(* IEC 61131-3 sources: moqui-plc/codesys-v4/moqui-plc.fbsdev/moqui.iecapp^/moqui/framework/src/main/org/moqui/mqtt, 4 files *)

(* ---- MqttConnectionFactory.fb.st ---- *)
(* Component to connect with a MQTT broker, using default configurations. *)
FUNCTION_BLOCK MqttConnectionFactory

	VAR_INPUT
		connect : BOOL := TRUE;
	END_VAR
	VAR_OUTPUT
		connection : MQTT.MQTTClient;
	    connected : BOOL;
	    busy : BOOL;
	    error : BOOL;
		errorId : INT;
	END_VAR
	VAR
		(* Connect properties v5 *)
		mqttConnectProperties : MQTT.MQTTConnectProperties := (
			udiSessionExpiryInterval := MoquiConf.sessionExpiryInterval,
			udiMaximumPacketSize := MoquiConf.maximumPacketSize
			(* userProperties := connectUserProperties *)
		);
		(* Will properties v5 *)
		mqttWillProperties : MQTT.MQTTWillProperties := (
			bPayloadFormatIndicator := MoquiConf.willPayloadFormatIndicator,
			udiMessageExpiryInterval := MoquiConf.willMessageExpiryInterval,
			wsContentType := MoquiConf.willContentType,
			udiWillDelayInterval := MoquiConf.willDelayInterval
			(* userProperties := willUserProperties *)
	    );
		(* TLS context *)
		cipherList : NBS.CIPHER_LIST := (psList := ADR('HIGH'), udiSize := 5);
		commonName : STRING := 'moqui';
	    certInfo : NBS.CERT_INFO := (psInfo := ADR(commonName), udiSize := INT_TO_UDINT(LEN(commonName)));
		defaultTlsContext : NBS.TLSContext := (
			sUseCaseName := commonName,
			ePurpose := NBS.PURPOSE.CLIENT_SIDE,
			sTLSVersion := '1.3',
			sCipherList := cipherList,
			sHostname := MoquiConf.brokerUrl,
			ciCertInfo := certInfo,
			udiVerificationMode	:= 2, (* 1 => No peer verification, 2 => Active Peer verification *)
			itfCertVerifer := 0
		);
		nullTlsContext : NBS.ITLSContext := 0;
		tlsContext : NBS.ITLSContext;
		useTLS : BOOL := FALSE;

		(*
	     * To use client certificates, configure the connection via the TLS context.
		 * Example:
		 *      commonName : STRING := 'COMMON_NAME_OF_CERTIFICATE'; // CN of the certificate (common name).
		 *      cipherList : NBS.CIPHER_LIST := (psList := ADR('HIGH'), udiSize := 5); // Cipher string see https://www.openssl.org/docs/man1.1.1/man1/ciphers.html
		 *      certInfo : NBS.CERT_INFO := (psInfo := ADR(commonName), udiSize := SIZEOF(commonName)); // CN of the certificate (common name)
		 *      tlsContext : NBS.TLSContext := (
		 *          sUseCaseName := commonName, // A certificate is stored in the certificate store with the use case name.
		 *          ePurpose := NBS.PURPOSE.CLIENT_SIDE, // For client certificates set this to NBS.PURPOSE.CLIENT_SIDE
	     *          sTLSVersion := '1.3', // The TLS version
	     *          sCipherList := cipherList, // Set the cipher list
	     *          sHostname := brokerUrl, // The hostname of the broker
	     *          udiVerificationMode := 2, // 2 => Active Peer verification
	     *          ciCertInfo := certInfo, // Set the cert info
	     *          itfCertVerifer := 0); // 0 => No Verifier
		 *      client : MQTT.MQTTClient := (itfTLSCOntext := _tlsContext);
		 * Use the method TLSContext.SetInitialValue to set the context while runtime and set the context via the input itfTLSCOntext of the client FB.
		 *)
	END_VAR

	(* TLS selection *)
	tlsContext := nullTlsContext;
	IF useTLS THEN tlsContext := defaultTlsContext; END_IF;

	(* Configure the MQTT connection *)
	connection(xEnable := connect, xConnectedToBroker => connected, xError => error, eMQTTerror => errorId,
		sHostname := MoquiConf.brokerUrl, uiPort := MoquiConf.brokerPort, sWebSocketUrl := MoquiConf.webSocketUrl, sClientId := MoquiConf.clientId,
		itfTLSContext := tlsContext, eCommunicationMode := MoquiConf.communicationMode, eMQTTVersion := MoquiConf.mqttVersion,
		wsUsername := MoquiConf.username, wsPassword := MoquiConf.password, mQTTConnectProperties := mqttConnectProperties,
		uiKeepAlive := MoquiConf.keepAlive, xCleanSession := MoquiConf.cleanSession, udiTimeOut := MoquiConf.timeout, tPingInterval := MoquiConf.pingInterval,
		wsWillTopic := MoquiConf.willTopic, pbWillMessage := ADR(MoquiConf.willMessage), uiWillMessageSize := INT_TO_UINT(LEN(MoquiConf.willMessage)),
		xWillRetain := MoquiConf.willRetain, eWillQoS := MoquiConf.willQoS, mQTTWillProperties := mqttWillProperties);
	END_FUNCTION_BLOCK

(* ---- MqttLogAppender.fb.st ---- *)
(*
 * Publishes one batch of log records as one MQTT message on logTopic.
 *
 * The broker connection belongs to MqttCommunication: this block only uses connectionFactory.connection.
 * A rising execute serializes the batch and publishes it; several steps run in the same call when they can.
 * done or error stay set until execute goes FALSE; then call the block until busy is FALSE before the next batch,
 * because the publisher and the JSON writer may still use the payload memory.
 *
 * errorId: 200 not connected to the broker; 100-113 serialization (SerializeLogToJson, serializeError = TRUE);
 * otherwise the MQTT error of the publisher (201 when the publisher reports an error without a code).
 *)
FUNCTION_BLOCK MqttLogAppender

	VAR_INPUT
	    execute : BOOL;
	    (* Data sources *)
	    logBuffer : REFERENCE TO ARRAY[1..MoquiConf.LOG_APPENDER_BATCH_SIZE] OF LogEvent;
	    logBufferSize : UINT;
	    (* The same batch was already sent once: set the DUP flag (QoS 1/2 only) *)
	    redelivery : BOOL;
	END_VAR
	VAR_OUTPUT
		done, busy, error : BOOL;
	    errorId : INT;
	    (* The error comes from the JSON serialization: a smaller batch may fit *)
	    serializeError : BOOL;
	END_VAR
	VAR
		state : MqttLogAppenderStatus := MqttLogAppenderStatus.Idle;
		finished : BOOL;
		pubTopic : WSTRING(1024) := MoquiConf.logTopic;
		(* Publisher *)
		publisher : MQTT.MQTTPublish;
		(* Publish properties v5 *)
		mqttPublishProperties : MQTT.MQTTPublishProperties := (
			bPayloadFormatIndicator := MoquiConf.pubPayloadFormatIndicator,
			wsContentType := MoquiConf.pubContentType,
			udiMessageExpiryInterval := MoquiConf.logMessageExpiryInterval
			(* userProperties := pubUserProperties *)
		);
	    (* JSON serializer *)
	    logMapper : SerializeLogToJson;
	END_VAR

	IF NOT execute THEN
		(* Release the JSON writer and the publisher; the payload stays untouched while either is busy *)
		logMapper(execute := FALSE);
		publisher(xExecute := FALSE, mqttClient := ec.connectionFactory.connection, wsTopicName := pubTopic);
		busy := logMapper.busy OR publisher.xBusy;
		done := FALSE;
		IF NOT busy THEN
			error := FALSE; errorId := 0; serializeError := FALSE;
			finished := FALSE;
			state := MqttLogAppenderStatus.Idle;
		END_IF;
		RETURN;
	END_IF;

	(* Outputs of the finished batch stay until execute goes FALSE *)
	IF finished THEN RETURN; END_IF;
	busy := TRUE;

	IF state = MqttLogAppenderStatus.Idle THEN
		IF NOT ec.connectionFactory.connected THEN
			error := TRUE; errorId := 200;
			busy := FALSE; finished := TRUE;
			RETURN;
		END_IF;
		state := MqttLogAppenderStatus.Serialize;
	END_IF;

	IF state = MqttLogAppenderStatus.Serialize THEN
		(* Compact output: no line breaks in the payload *)
		logMapper(execute := TRUE, logBuffer := logBuffer, logBufferSize := logBufferSize, lineBreak := "");
		IF logMapper.error THEN
			error := TRUE; errorId := logMapper.errorId; serializeError := TRUE;
			busy := FALSE; finished := TRUE;
			RETURN;
		ELSIF logMapper.done THEN
			state := MqttLogAppenderStatus.Publish;
		END_IF;
	END_IF;

	IF state = MqttLogAppenderStatus.Publish THEN
		publisher(xExecute := TRUE, mqttClient := ec.connectionFactory.connection, wsTopicName := pubTopic,
			pbPayload := ADR(logMapper.jsonPayload), udiPayloadSize := logMapper.payloadSize,
			eQoS := MoquiConf.logPubQoS, xReDelivery := redelivery AND (MoquiConf.logPubQoS <> MQTT.MQTT_QOS.QoS0),
			xRetain := MoquiConf.logPubRetain, udiTimeOut := MoquiConf.logAppenderTimeout,
			mQTTPublishProperties := mqttPublishProperties);
		IF publisher.xError THEN
			error := TRUE; errorId := TO_INT(publisher.eMQTTError);
			IF errorId = 0 THEN errorId := 201; END_IF;
			busy := FALSE; finished := TRUE;
		ELSIF publisher.xDone THEN
			done := TRUE;
			busy := FALSE; finished := TRUE;
		END_IF;
	END_IF;
	END_FUNCTION_BLOCK

(* ---- MqttParameterPub.prg.st ---- *)
(*
 * Optional publisher for parameter replication between peer PLCs/Applications,
 * typically for a developer-defined redundancy strategy. Operational numeric
 * and textual telemetry is published by LogDispatcher instead.
 * Called by MqttCommunication, which owns the broker connection.
 *)
PROGRAM MqttParameterPub

	VAR
		done, busy, error : BOOL;
	    errorId : INT;
		jsonPayload : WSTRING(MoquiConf.JSON_PAYLOAD_MAX_SIZE);
		pubTopic : WSTRING(1024) := MoquiConf.liveParamsPubTopic;
		pubMessage : STRING(MoquiConf.JSON_PAYLOAD_MAX_SIZE);
		(* Publisher *)
		publisher : MQTT.MQTTPublish;
		(* Publish properties v5 *)
		mqttPublishProperties : MQTT.MQTTPublishProperties := (
			bPayloadFormatIndicator := MoquiConf.pubPayloadFormatIndicator,
			wsContentType := MoquiConf.pubContentType,
			udiMessageExpiryInterval := MoquiConf.pubMessageExpiryInterval
			(* userProperties := pubUserProperties *)
		);
	    (* JSON serializer *)
	    parameterMapper : SerializeParametersToJson;
	END_VAR

	(* Publishing disabled *)
	IF NOT ec.paramsPubEnable THEN
		parameterMapper(execute := FALSE);
		publisher(xExecute := FALSE, mqttClient := ec.connectionFactory.connection, wsTopicName := pubTopic);
		done := FALSE; busy := FALSE; error := FALSE; errorId := 0;
		RETURN;
	END_IF;

	(* Waiting for connection to broker *)
	IF NOT ec.connectionFactory.connected THEN RETURN; END_IF;

	IF NOT publisher.xBusy THEN
		(* JSON mapping *)
		parameterMapper(execute := TRUE, jsonPayload => jsonPayload,
			busy => busy, error => error, errorId => errorId);
		IF parameterMapper.error THEN
			(* Reset JSON writer *)
			parameterMapper(execute := FALSE, error => error, errorId => errorId);
			done := FALSE; busy := FALSE;
			RETURN;
		END_IF;
	END_IF;

	IF parameterMapper.done THEN
		(* Publish the payload *)
		pubMessage := TO_STRING(jsonPayload);
		publisher(xExecute := TRUE, mqttClient := ec.connectionFactory.connection, wsTopicName := pubTopic,
			pbPayload := ADR(pubMessage), udiPayloadSize := INT_TO_UDINT(LEN(pubMessage)),
			eQoS := MoquiConf.paramsPubQoS, xReDelivery := MoquiConf.paramsReDelivery, xRetain := MoquiConf.paramsPubRetain,
			udiTimeOut := MoquiConf.liveParamsPubTimeout, mQTTPublishProperties := mqttPublishProperties,
			xDone => done, xBusy => busy, xError => error, eMQTTError => errorId);

		IF publisher.xError OR publisher.xDone THEN
			(* Auto reset: next cycle restarts from scratch *)
			parameterMapper(execute := FALSE, busy => busy,
				error => error, errorId => errorId);
			publisher(xExecute := FALSE, mqttClient := ec.connectionFactory.connection, wsTopicName := pubTopic,
				xDone => done, xBusy => busy, xError => error, eMQTTError => errorId);
		END_IF;
	END_IF;
	END_PROGRAM

(* ---- MqttParameterSub.prg.st ---- *)
(*
 * Live parameter writes from Moqui: subscribes liveParamsSubTopic and applies each payload with
 * DeserializeJsonToParameters. Called by MqttCommunication, which owns the broker connection.
 *)
PROGRAM MqttParameterSub

	VAR
		done, busy, error : BOOL;
	    errorId : INT;
		(* Subscriber *)
		subscriber : MQTT.MQTTSubscribe;
		(* Subscribe properties v5 *)
		mqttSubscribeProperties : MQTT.MQTTSubscribeProperties := (
			udiSubscriptionIdentifier := MoquiConf.subscriptionIdentifier,
			xNoLocalOption := MoquiConf.subNoLocalOption,
			xRetainAsPublished := MoquiConf.subRetainAsPublished,
			eRetainHandling := MoquiConf.subRetainHandling
			(* userProperties := subUserProperties; *)
		);
	    (* JSON parser *)
	    parser : DeserializeJsonToParameters;
		parserActive : BOOL; (* TRUE while parser is running across multiple cycles *)
		subTopicFilter : WSTRING(1024) := MoquiConf.liveParamsSubTopic;
		(* Last incoming message *)
		rxBuffer : STRING(MoquiConf.JSON_PAYLOAD_MAX_SIZE);
		pRxBytes : POINTER TO ARRAY[0..MoquiConf.JSON_PAYLOAD_MAX_SIZE] OF BYTE;
		clearIdx : UINT;
		lastSubMessage : STRING(MoquiConf.JSON_PAYLOAD_MAX_SIZE);
	    receivedPayload : WSTRING(MoquiConf.JSON_PAYLOAD_MAX_SIZE);
		subscriberEnable : BOOL;
	END_VAR

	(* Subscription disabled *)
	IF NOT ec.paramsSubEnable THEN
		subscriber(xEnable := FALSE, mqttClient := ec.connectionFactory.connection, wsTopicFilter := subTopicFilter);
		parser(execute := FALSE);
		parserActive := FALSE;
		done := FALSE; busy := FALSE; error := FALSE; errorId := 0;
	    RETURN;
	END_IF;

	(* Manage subscriber enable: disable for one cycle on error to reset the FB *)
	IF subscriber.xError THEN
		subscriberEnable := FALSE;
	ELSE
		subscriberEnable := ec.connectionFactory.connected;
	END_IF;

	(* Drive subscriber continuously; xDone = subscription confirmed (sub ack), not end of session *)
	subscriber(xEnable := subscriberEnable, mqttClient := ec.connectionFactory.connection,
		eFilterMode := MoquiConf.paramsSubFilterMode, wsTopicFilter := subTopicFilter, eSubscribeQoS := MoquiConf.paramsSubQoS,
		udiTimeout := MoquiConf.liveParamsSubTimeout, pbPayload := ADR(rxBuffer),
		udiMaxPayloadSize := SIZEOF(rxBuffer) - 1, mQTTSubscribeProperties := mqttSubscribeProperties,
		xDone => done, xBusy => busy, xError => error, eMQTTError => errorId);

	(* xReceived pulses TRUE for one cycle only: copy NUL-terminated buffer, clear rxBuffer, and latch parserActive *)
	IF subscriber.xReceived THEN
		IF subscriber.xSubscribeActive AND subscriber.wsLastTopic = subTopicFilter THEN
			lastSubMessage := rxBuffer;
			receivedPayload := TO_WSTRING(lastSubMessage);
			IF parserActive THEN
				parser(execute := FALSE);
			END_IF;
			parserActive := TRUE;
		END_IF;
		pRxBytes := ADR(rxBuffer);
		FOR clearIdx := 0 TO MoquiConf.JSON_PAYLOAD_MAX_SIZE DO
			IF pRxBytes^[clearIdx] = 0 THEN
				EXIT;
			END_IF;
			pRxBytes^[clearIdx] := 0;
		END_FOR;
	END_IF;

	(* Drive parser every cycle until done/error, regardless of xReceived *)
	IF parserActive THEN
		(* JSON parsing *)
		parser(execute := TRUE, jsonPayload := receivedPayload,
			busy => busy, error => error, errorId => errorId);

		IF parser.done OR parser.error THEN
			(* Auto reset: next cycle restarts from scratch *)
			parser(execute := FALSE, done => done, busy => busy,
				error => error, errorId => errorId);
			parserActive := FALSE;
		END_IF;
	END_IF;
	END_PROGRAM
